// TIA Portal V19 export
VAR_GLOBAL   // PLC tag table "Test"
END_VAR
